Yaskawa INFORM job: CHAMFER.JBI

/JOB
//NAME CHAMFER
//POS
///NPOS 111,0,0,0,0,0
///TOOL 9
///POSTYPE PULSE
///PULSE
C00000=-44,20,38,3,-108,94
C00001=-44,20,38,3,-108,94
C00002=-37,19,37,3,-107,87
C00003=-37,19,37,3,-107,87
C00004=-37,19,34,4,-105,88
C00005=-37,17,30,3,-103,87
C00006=-38,16,27,2,-101,87
C00007=-38,15,24,1,-98,87
C00008=-38,14,21,0,-96,87
C00009=-38,13,18,-1,-94,87
C00010=-38,13,15,-2,-92,87
C00011=-39,13,13,-2,-90,88
C00012=-39,12,10,-4,-88,86
C00013=-39,12,9,-3,-87,88
C00014=-39,12,9,-3,-87,88
C00015=-38,12,9,-2,-86,88
C00016=-38,12,9,0,-86,87
C00017=-37,12,9,3,-87,85
C00018=-37,12,9,6,-87,84
C00019=-36,13,9,8,-87,83
C00020=-36,13,9,10,-87,81
C00021=-35,13,9,12,-88,80
C00022=-35,14,10,15,-89,78
C00023=-34,14,10,17,-90,76
C00024=-34,14,10,20,-91,74
C00025=-33,15,11,21,-92,72
C00026=-33,15,11,23,-94,69
C00027=-33,16,12,25,-96,66
C00028=-32,17,12,26,-98,64
C00029=-32,17,13,27,-101,61
C00030=-32,18,14,28,-104,58
C00031=-32,19,14,28,-106,55
C00032=-32,19,15,27,-109,51
C00033=-32,20,16,26,-111,47
C00034=-32,21,17,24,-114,42
C00035=-33,21,17,22,-115,39
C00036=-33,21,18,20,-117,34
C00037=-33,21,18,18,-117,30
C00038=-34,21,18,15,-118,26
C00039=-34,21,18,12,-117,21
C00040=-34,21,17,9,-116,17
C00041=-35,20,16,7,-115,13
C00042=-35,19,16,5,-113,9
C00043=-35,19,16,4,-112,8
C00044=-36,18,15,3,-109,5
C00045=-36,17,14,2,-107,3
C00046=-36,17,13,1,-104,1
C00047=-36,16,12,0,-102,0
C00048=-36,15,11,0,-99,-2
C00049=-36,14,11,0,-97,-2
C00050=-36,13,10,0,-95,-3
C00051=-37,13,9,0,-92,-4
C00052=-37,12,8,0,-89,-4
C00053=-37,11,7,0,-86,-5
C00054=-37,10,7,1,-85,-5
C00055=-37,10,7,1,-84,-5
C00056=-37,10,7,1,-84,-5
C00057=-36,10,8,1,-85,-6
C00058=-37,10,11,1,-88,-4
C00059=-37,11,13,1,-91,-4
C00060=-37,12,16,0,-94,-4
C00061=-37,13,19,0,-96,-4
C00062=-37,14,22,0,-99,-5
C00063=-37,15,26,0,-102,-4
C00064=-37,16,29,0,-105,-5
C00065=-37,18,34,0,-109,-3
C00066=-37,19,36,0,-110,-4
C00067=-37,19,36,0,-110,-4
C00068=-37,19,38,0,-111,-5
C00069=-37,18,36,0,-108,-5
C00070=-36,17,35,1,-105,-4
C00071=-36,16,33,1,-102,-4
C00072=-36,15,32,1,-99,-3
C00073=-36,14,31,1,-96,-2
C00074=-36,13,30,1,-94,-2
C00075=-36,12,28,1,-91,0
C00076=-36,11,26,0,-88,1
C00077=-36,10,25,-1,-84,3
C00078=-36,9,24,-2,-82,5
C00079=-37,8,22,-3,-79,8
C00080=-37,7,21,-5,-76,11
C00081=-38,7,20,-7,-75,14
C00082=-38,6,19,-9,-73,19
C00083=-39,6,18,-12,-72,24
C00084=-40,6,17,-15,-71,28
C00085=-40,6,17,-18,-71,34
C00086=-41,7,18,-22,-72,39
C00087=-42,7,19,-25,-74,45
C00088=-42,8,19,-27,-76,49
C00089=-43,9,21,-28,-79,54
C00090=-43,10,22,-29,-82,57
C00091=-44,12,24,-30,-85,61
C00092=-44,13,26,-30,-89,64
C00093=-44,15,29,-29,-92,67
C00094=-44,16,31,-28,-95,70
C00095=-43,17,33,-26,-98,72
C00096=-43,17,33,-25,-99,73
C00097=-43,18,35,-23,-101,75
C00098=-42,19,36,-21,-103,77
C00099=-42,20,38,-18,-105,79
C00100=-41,20,39,-16,-106,81
C00101=-41,21,40,-13,-107,82
C00102=-40,21,39,-11,-108,83
C00103=-40,20,39,-9,-108,84
C00104=-39,20,39,-6,-108,85
C00105=-38,20,39,-3,-108,86
C00106=-38,20,39,0,-108,87
C00107=-37,20,38,2,-108,87
C00108=-37,19,37,3,-107,87
C00109=-37,19,37,3,-107,87
C00110=-44,20,38,3,-108,94
//INST
///DATE 2026/10/26 01:19
///COMM Generated using RoboDK
///ATTR SC,RW
///GROUP1 RB1
NOP
'Program generated by Vertical
'Bot Studio for Motoman ES200D
' on 25/10/2026 12:00:00
'Using nominal kinematics.
'Using Frame 1 (targets wrt ba
'se):
'1724.5,-1789.7,1123.6,0.0,0.0
',93.8
'Tool Spindle should be close
'to:
'417.9,0.0,132.0,0.0,90.0,0.0
CALL JOB:ONCHAMF
'Using Frame 1 (targets wrt ba
'se):
'1724.5,-1789.7,1123.6,0.0,0.0
',93.8
'Tool Spindle should be close
'to:
'417.9,0.0,132.0,0.0,90.0,0.0
'show Spindle
MOVJ C00000 VJ=50.00
CALL JOB:ONCHAMF
MOVL C00001 V=1000.0
MOVL C00002 V=1000.0
CALL JOB:ONCHAMF
MOVL C00003 V=1000.0
MOVL C00004 V=50.0
MOVL C00005 V=50.0
MOVL C00006 V=50.0
MOVL C00007 V=50.0
MOVL C00008 V=50.0
MOVL C00009 V=50.0
MOVL C00010 V=50.0
MOVL C00011 V=50.0
MOVL C00012 V=50.0
MOVL C00013 V=50.0
MOVL C00014 V=50.0
MOVL C00015 V=50.0
MOVL C00016 V=50.0
MOVL C00017 V=50.0
MOVL C00018 V=50.0
MOVL C00019 V=50.0
MOVL C00020 V=50.0
MOVL C00021 V=50.0
MOVL C00022 V=50.0
MOVL C00023 V=50.0
MOVL C00024 V=50.0
MOVL C00025 V=50.0
MOVL C00026 V=50.0
MOVL C00027 V=50.0
MOVL C00028 V=50.0
MOVL C00029 V=50.0
MOVL C00030 V=50.0
MOVL C00031 V=50.0
MOVL C00032 V=50.0
MOVL C00033 V=50.0
MOVL C00034 V=50.0
MOVL C00035 V=50.0
MOVL C00036 V=50.0
MOVL C00037 V=50.0
MOVL C00038 V=50.0
MOVL C00039 V=50.0
MOVL C00040 V=50.0
MOVL C00041 V=50.0
MOVL C00042 V=50.0
MOVL C00043 V=50.0
MOVL C00044 V=50.0
MOVL C00045 V=50.0
MOVL C00046 V=50.0
MOVL C00047 V=50.0
MOVL C00048 V=50.0
MOVL C00049 V=50.0
MOVL C00050 V=50.0
MOVL C00051 V=50.0
MOVL C00052 V=50.0
MOVL C00053 V=50.0
MOVL C00054 V=50.0
MOVL C00055 V=50.0
MOVL C00056 V=50.0
MOVL C00057 V=50.0
MOVL C00058 V=50.0
MOVL C00059 V=50.0
MOVL C00060 V=50.0
MOVL C00061 V=50.0
MOVL C00062 V=50.0
MOVL C00063 V=50.0
MOVL C00064 V=50.0
MOVL C00065 V=50.0
MOVL C00066 V=50.0
MOVL C00067 V=50.0
MOVL C00068 V=50.0
MOVL C00069 V=50.0
MOVL C00070 V=50.0
MOVL C00071 V=50.0
MOVL C00072 V=50.0
MOVL C00073 V=50.0
MOVL C00074 V=50.0
MOVL C00075 V=50.0
MOVL C00076 V=50.0
MOVL C00077 V=50.0
MOVL C00078 V=50.0
MOVL C00079 V=50.0
MOVL C00080 V=50.0
MOVL C00081 V=50.0
MOVL C00082 V=50.0
MOVL C00083 V=50.0
MOVL C00084 V=50.0
MOVL C00085 V=50.0
MOVL C00086 V=50.0
MOVL C00087 V=50.0
MOVL C00088 V=50.0
MOVL C00089 V=50.0
MOVL C00090 V=50.0
MOVL C00091 V=50.0
MOVL C00092 V=50.0
MOVL C00093 V=50.0
MOVL C00094 V=50.0
MOVL C00095 V=50.0
MOVL C00096 V=50.0
MOVL C00097 V=50.0
MOVL C00098 V=50.0
MOVL C00099 V=50.0
MOVL C00100 V=50.0
MOVL C00101 V=50.0
MOVL C00102 V=50.0
MOVL C00103 V=50.0
MOVL C00104 V=50.0
MOVL C00105 V=50.0
MOVL C00106 V=50.0
MOVL C00107 V=50.0
MOVL C00108 V=50.0
CALL JOB:ONCHAMF
MOVL C00109 V=1000.0
MOVL C00110 V=1000.0
CALL JOB:ONCHAMF
END
